(* IEC 61131-3 sources: SortJet_MasterSPS_Aufbau.fbsproj/Device.device.xml.v3^/Plc Logic.plclogic.xml.v3^/Application.application.xml.v3^/09_Station/Stationen/Faecherwagen [301-305]/0_Konfig, 5 files *)

(* ---- MK_Faecherwagen.gvl ---- *)
(* METADATA
{
	"v3Meta": {
		"objectGuid": "4f007b85-dd1b-4818-92fb-7451563e5cb0"
	}
}
*)
{attribute 'allow_unqualified_access'}
NAMESPACE MK_Faecherwagen
VAR_GLOBAL
  apgMKFaecherwagenstation : ARRAY[cERSTE_FAECHERWAGENSTATIONS_NR..cLETZTE_FAECHERWAGENSTATIONS_NR] OF Parameter_Station :=[
    (
     stStationsNummern         := (  NummerIntern    :=   301,                                 // Stationsnummer fuer das MMI und die Stationsangabe der Meldungen
                                     NummerExtern    :=  1301,                                 // Stationsnummer fuer Bedienermeldungen
                                     NummerSPS       :=   301 ),                               // Stationsnummer SPS-intern (Indizes)
      bDeaktivieren             := FALSE,                                                      // Station deaktiviert (keine Auftraege, keine Referenzfahrt)
      wMeldungsNummer           := 1400,                                                       // Basis-Meldungsnummer (WatchIO)
      eStationsTyp              := eFaecherwagen,                                              // Typ der Station
      eaAutomatikkreis          := [eAutomatikkreis_2],                                        // Automatikkreise, zu denen die Station gehoert
     // stStationsParameter
     // stSchnittstellendaten
     // stFremdanlage
     // stGlasdaten
      eaSicherheitskreis        := [eSicherheitskreis_1],                                      // Sicherheitskreise, in die die Station eingebunden ist
      // astSicherheitskreisTeilabschaltung
      eSystemcheckZyklus        := eSystemcheckZyklus_1,                                       // In welchem Zyklus des Systemchecks die Station geprueft wird
     // stStationsOptionen
      stStationsAufbau          := ( bAnschlag                     := FALSE,                   // Ausbaustufe: Ausrichtanschlaege
                                     bRolltor                      := TRUE,                    // Ausbaustufe Faecherwagen: Rolltor
                                     bKlemmzylinder                := FALSE,                   // Ausbaustufe Faecherwagen: Klemmzylinder fixiert den Oberrahmen beim Ein- und Ausschleusen
                                     bGreifer                      := [cANZAHL_WAENDE(FALSE)], // Shuttle: Greifer je Wand (Scheibe aus dem Faecherwagen ziehen bzw. hineinschieben)
                                     bRFID                         := TRUE,                    // RFID-Leser vorhanden
                                     bAGV                          := FALSE,                   // Ausbaustufe Faecherwagen: Betrieb mit AGV
                                     bGeblase                      := [ FALSE ],               // Ausbaustufe: Geblaese je Wand
                                     bGlastransport                := [ FALSE ],               // Ausbaustufe: Glastransport je Wand
                                     bKippen                       := [ FALSE ],               // Ausbaustufe: Kippen je Wand
                                     bTransportVerstellung         := [ FALSE ],               // Ausbaustufe Shuttle: Transport-/Dickenverstellung je Wand
                                     bWandverstellung              := [ FALSE ],               // Ausbaustufe Station: Wandverstellung je Wand
                                     bWandverstellungMotorisch     := FALSE,                   // Shuttle: Transport-/Wandverstellung mit Antrieb statt pneumatisch
                                     bRoellchenleiste              := [ FALSE ],               // Ausbaustufe Station: Roellchenleiste je Wand
                                     bHub                          := FALSE,                   // Ausbaustufe: Hub der Station
                                     bHubrahmen                    := FALSE,                   // Ausbaustufe: Hubrahmen (Riemen heben/senken)
                                     bDrehen                       := FALSE,                   // Ausbaustufe: Drehen
                                     bQuerachse                    := FALSE,                   // Ausbaustufe: Querachse
                                     bMessachse                    := FALSE,                   // Ausbaustufe: Messachse (Anlegetisch, Anlegewand)
                                     bDruckluft                    := FALSE,                   // Druckluftueberwachung vorhanden
                                     bSensorAuslauf                := FALSE,                   // Auslaufsensor vorhanden
                                     bSensorEinlauf                := FALSE,                   // Einlaufsensor vorhanden
                                     bSensorEinlaufStopp           := FALSE,                   // Shuttle: zusaetzlicher Stopp-Sensor am Einlauf (ohne: Einlaufsensor), Gegenstueck zum Auslauf-Stopp im Rueckwaertstransport
                                     bSensorAuslaufStopp           := FALSE,                   // Shuttle: zusaetzlicher Stopp-Sensor am Auslauf (ohne: Auslaufsensor), Verfahrfreigabe und Scheibe hat Shuttle verlassen
                                     bDurchlaufSperreZumNachfolger := FALSE,                   // Ausbaustufe: bewegliche Abschrankung zum Nachfolger
                                     bKippenSchuetz                := FALSE,                   // Kippen ueber Schuetz statt Umrichter
                                     bQuerfahrt                    := FALSE,                   // Ausbaustufe: Querfahrt
                                     bDurchgang                    := FALSE,                   // Station ist Teil eines Durchgangs (belegt = Oeffnen blockiert)
                                     bSlaveAntrieb                 := FALSE,                   // Glastransport mit Slave-Antrieb
                                     bKipparme                     := FALSE,                   // Ausbaustufe: Kipparme
                                     bMessachseAmEndeVomTisch      := FALSE,                   // Messachse am Ende des Tisches (Hoehenfehler fragt den Bediener)
                                     bDLSSchmiersystem             := FALSE,                   // Zentralschmierung DLS vorhanden
                                     bGlastransportSlaveVorhanden  := FALSE,                   // Glastransport mit Slave-Antrieb (Meldungen/Ueberwachung Slave)
                                     wHydraulikstation             := cHYDRAULIKSTATION_1      // Faecherwagen Hydraulik: zugeordnete Hydraulikstation (cHYDRAULIKSTATION_x), 0 = keine
                                    )
     // astShuttleAnhaltenQuellen
    ),
    (
     stStationsNummern         := (  NummerIntern    :=   302,                                 // Stationsnummer fuer das MMI und die Stationsangabe der Meldungen
                                     NummerExtern    :=  1302,                                 // Stationsnummer fuer Bedienermeldungen
                                     NummerSPS       :=   302 ),                               // Stationsnummer SPS-intern (Indizes)
      bDeaktivieren             := FALSE,                                                      // Station deaktiviert (keine Auftraege, keine Referenzfahrt)
      wMeldungsNummer           := 1420,                                                       // Basis-Meldungsnummer (WatchIO)
      eStationsTyp              := eFaecherwagen,                                              // Typ der Station
      eaAutomatikkreis          := [eAutomatikkreis_2],                                        // Automatikkreise, zu denen die Station gehoert
     // stStationsParameter
     // stSchnittstellendaten
     // stFremdanlage
     // stGlasdaten
      eaSicherheitskreis        := [eSicherheitskreis_1],                                      // Sicherheitskreise, in die die Station eingebunden ist
      // astSicherheitskreisTeilabschaltung
      eSystemcheckZyklus        := eSystemcheckZyklus_1,                                       // In welchem Zyklus des Systemchecks die Station geprueft wird
     // stStationsOptionen
      stStationsAufbau          := ( bAnschlag                     := FALSE,                   // Ausbaustufe: Ausrichtanschlaege
                                     bRolltor                      := TRUE,                    // Ausbaustufe Faecherwagen: Rolltor
                                     bKlemmzylinder                := FALSE,                   // Ausbaustufe Faecherwagen: Klemmzylinder fixiert den Oberrahmen beim Ein- und Ausschleusen
                                     bGreifer                      := [cANZAHL_WAENDE(FALSE)], // Shuttle: Greifer je Wand (Scheibe aus dem Faecherwagen ziehen bzw. hineinschieben)
                                     bRFID                         := TRUE,                    // RFID-Leser vorhanden
                                     bAGV                          := FALSE,                   // Ausbaustufe Faecherwagen: Betrieb mit AGV
                                     bGeblase                      := [ FALSE ],               // Ausbaustufe: Geblaese je Wand
                                     bGlastransport                := [ FALSE ],               // Ausbaustufe: Glastransport je Wand
                                     bKippen                       := [ FALSE ],               // Ausbaustufe: Kippen je Wand
                                     bTransportVerstellung         := [ FALSE ],               // Ausbaustufe Shuttle: Transport-/Dickenverstellung je Wand
                                     bWandverstellung              := [ FALSE ],               // Ausbaustufe Station: Wandverstellung je Wand
                                     bWandverstellungMotorisch     := FALSE,                   // Shuttle: Transport-/Wandverstellung mit Antrieb statt pneumatisch
                                     bRoellchenleiste              := [ FALSE ],               // Ausbaustufe Station: Roellchenleiste je Wand
                                     bHub                          := FALSE,                   // Ausbaustufe: Hub der Station
                                     bHubrahmen                    := FALSE,                   // Ausbaustufe: Hubrahmen (Riemen heben/senken)
                                     bDrehen                       := FALSE,                   // Ausbaustufe: Drehen
                                     bQuerachse                    := FALSE,                   // Ausbaustufe: Querachse
                                     bMessachse                    := FALSE,                   // Ausbaustufe: Messachse (Anlegetisch, Anlegewand)
                                     bDruckluft                    := FALSE,                   // Druckluftueberwachung vorhanden
                                     bSensorAuslauf                := FALSE,                   // Auslaufsensor vorhanden
                                     bSensorEinlauf                := FALSE,                   // Einlaufsensor vorhanden
                                     bSensorEinlaufStopp           := FALSE,                   // Shuttle: zusaetzlicher Stopp-Sensor am Einlauf (ohne: Einlaufsensor), Gegenstueck zum Auslauf-Stopp im Rueckwaertstransport
                                     bSensorAuslaufStopp           := FALSE,                   // Shuttle: zusaetzlicher Stopp-Sensor am Auslauf (ohne: Auslaufsensor), Verfahrfreigabe und Scheibe hat Shuttle verlassen
                                     bDurchlaufSperreZumNachfolger := FALSE,                   // Ausbaustufe: bewegliche Abschrankung zum Nachfolger
                                     bKippenSchuetz                := FALSE,                   // Kippen ueber Schuetz statt Umrichter
                                     bQuerfahrt                    := FALSE,                   // Ausbaustufe: Querfahrt
                                     bDurchgang                    := FALSE,                   // Station ist Teil eines Durchgangs (belegt = Oeffnen blockiert)
                                     bSlaveAntrieb                 := FALSE,                   // Glastransport mit Slave-Antrieb
                                     bKipparme                     := FALSE,                   // Ausbaustufe: Kipparme
                                     bMessachseAmEndeVomTisch      := FALSE,                   // Messachse am Ende des Tisches (Hoehenfehler fragt den Bediener)
                                     bDLSSchmiersystem             := FALSE,                   // Zentralschmierung DLS vorhanden
                                     bGlastransportSlaveVorhanden  := FALSE,                   // Glastransport mit Slave-Antrieb (Meldungen/Ueberwachung Slave)
                                     wHydraulikstation             := cHYDRAULIKSTATION_1      // Faecherwagen Hydraulik: zugeordnete Hydraulikstation (cHYDRAULIKSTATION_x), 0 = keine
                                    )
     // astShuttleAnhaltenQuellen
    ),
    (
     stStationsNummern         := (  NummerIntern    :=   303,                                 // Stationsnummer fuer das MMI und die Stationsangabe der Meldungen
                                     NummerExtern    :=  1303,                                 // Stationsnummer fuer Bedienermeldungen
                                     NummerSPS       :=   303 ),                               // Stationsnummer SPS-intern (Indizes)
      bDeaktivieren             := FALSE,                                                      // Station deaktiviert (keine Auftraege, keine Referenzfahrt)
      wMeldungsNummer           := 1440,                                                       // Basis-Meldungsnummer (WatchIO)
      eStationsTyp              := eFaecherwagen,                                              // Typ der Station
      eaAutomatikkreis          := [eAutomatikkreis_2],                                        // Automatikkreise, zu denen die Station gehoert
     // stStationsParameter
     // stSchnittstellendaten
     // stFremdanlage
     // stGlasdaten
      eaSicherheitskreis        := [eSicherheitskreis_1],                                      // Sicherheitskreise, in die die Station eingebunden ist
      // astSicherheitskreisTeilabschaltung
      eSystemcheckZyklus        := eSystemcheckZyklus_1,                                       // In welchem Zyklus des Systemchecks die Station geprueft wird
     // stStationsOptionen
      stStationsAufbau          := ( bAnschlag                     := FALSE,                   // Ausbaustufe: Ausrichtanschlaege
                                     bRolltor                      := TRUE,                    // Ausbaustufe Faecherwagen: Rolltor
                                     bKlemmzylinder                := FALSE,                   // Ausbaustufe Faecherwagen: Klemmzylinder fixiert den Oberrahmen beim Ein- und Ausschleusen
                                     bGreifer                      := [cANZAHL_WAENDE(FALSE)], // Shuttle: Greifer je Wand (Scheibe aus dem Faecherwagen ziehen bzw. hineinschieben)
                                     bRFID                         := TRUE,                    // RFID-Leser vorhanden
                                     bAGV                          := FALSE,                   // Ausbaustufe Faecherwagen: Betrieb mit AGV
                                     bGeblase                      := [ FALSE ],               // Ausbaustufe: Geblaese je Wand
                                     bGlastransport                := [ FALSE ],               // Ausbaustufe: Glastransport je Wand
                                     bKippen                       := [ FALSE ],               // Ausbaustufe: Kippen je Wand
                                     bTransportVerstellung         := [ FALSE ],               // Ausbaustufe Shuttle: Transport-/Dickenverstellung je Wand
                                     bWandverstellung              := [ FALSE ],               // Ausbaustufe Station: Wandverstellung je Wand
                                     bWandverstellungMotorisch     := FALSE,                   // Shuttle: Transport-/Wandverstellung mit Antrieb statt pneumatisch
                                     bRoellchenleiste              := [ FALSE ],               // Ausbaustufe Station: Roellchenleiste je Wand
                                     bHub                          := FALSE,                   // Ausbaustufe: Hub der Station
                                     bHubrahmen                    := FALSE,                   // Ausbaustufe: Hubrahmen (Riemen heben/senken)
                                     bDrehen                       := FALSE,                   // Ausbaustufe: Drehen
                                     bQuerachse                    := FALSE,                   // Ausbaustufe: Querachse
                                     bMessachse                    := FALSE,                   // Ausbaustufe: Messachse (Anlegetisch, Anlegewand)
                                     bDruckluft                    := FALSE,                   // Druckluftueberwachung vorhanden
                                     bSensorAuslauf                := FALSE,                   // Auslaufsensor vorhanden
                                     bSensorEinlauf                := FALSE,                   // Einlaufsensor vorhanden
                                     bSensorEinlaufStopp           := FALSE,                   // Shuttle: zusaetzlicher Stopp-Sensor am Einlauf (ohne: Einlaufsensor), Gegenstueck zum Auslauf-Stopp im Rueckwaertstransport
                                     bSensorAuslaufStopp           := FALSE,                   // Shuttle: zusaetzlicher Stopp-Sensor am Auslauf (ohne: Auslaufsensor), Verfahrfreigabe und Scheibe hat Shuttle verlassen
                                     bDurchlaufSperreZumNachfolger := FALSE,                   // Ausbaustufe: bewegliche Abschrankung zum Nachfolger
                                     bKippenSchuetz                := FALSE,                   // Kippen ueber Schuetz statt Umrichter
                                     bQuerfahrt                    := FALSE,                   // Ausbaustufe: Querfahrt
                                     bDurchgang                    := FALSE,                   // Station ist Teil eines Durchgangs (belegt = Oeffnen blockiert)
                                     bSlaveAntrieb                 := FALSE,                   // Glastransport mit Slave-Antrieb
                                     bKipparme                     := FALSE,                   // Ausbaustufe: Kipparme
                                     bMessachseAmEndeVomTisch      := FALSE,                   // Messachse am Ende des Tisches (Hoehenfehler fragt den Bediener)
                                     bDLSSchmiersystem             := FALSE,                   // Zentralschmierung DLS vorhanden
                                     bGlastransportSlaveVorhanden  := FALSE,                   // Glastransport mit Slave-Antrieb (Meldungen/Ueberwachung Slave)
                                     wHydraulikstation             := cHYDRAULIKSTATION_1      // Faecherwagen Hydraulik: zugeordnete Hydraulikstation (cHYDRAULIKSTATION_x), 0 = keine
                                    )
     // astShuttleAnhaltenQuellen
    ),
    (
     stStationsNummern         := (  NummerIntern    :=   304,                                 // Stationsnummer fuer das MMI und die Stationsangabe der Meldungen
                                     NummerExtern    :=  1304,                                 // Stationsnummer fuer Bedienermeldungen
                                     NummerSPS       :=   304 ),                               // Stationsnummer SPS-intern (Indizes)
      bDeaktivieren             := FALSE,                                                      // Station deaktiviert (keine Auftraege, keine Referenzfahrt)
      wMeldungsNummer           := 1460,                                                       // Basis-Meldungsnummer (WatchIO)
      eStationsTyp              := eFaecherwagen,                                              // Typ der Station
      eaAutomatikkreis          := [eAutomatikkreis_2],                                        // Automatikkreise, zu denen die Station gehoert
     // stStationsParameter
     // stSchnittstellendaten
     // stFremdanlage
     // stGlasdaten
      eaSicherheitskreis        := [eSicherheitskreis_1],                                      // Sicherheitskreise, in die die Station eingebunden ist
      // astSicherheitskreisTeilabschaltung
      eSystemcheckZyklus        := eSystemcheckZyklus_1,                                       // In welchem Zyklus des Systemchecks die Station geprueft wird
     // stStationsOptionen
      stStationsAufbau          := ( bAnschlag                     := FALSE,                   // Ausbaustufe: Ausrichtanschlaege
                                     bRolltor                      := TRUE,                    // Ausbaustufe Faecherwagen: Rolltor
                                     bKlemmzylinder                := FALSE,                   // Ausbaustufe Faecherwagen: Klemmzylinder fixiert den Oberrahmen beim Ein- und Ausschleusen
                                     bGreifer                      := [cANZAHL_WAENDE(FALSE)], // Shuttle: Greifer je Wand (Scheibe aus dem Faecherwagen ziehen bzw. hineinschieben)
                                     bRFID                         := TRUE,                    // RFID-Leser vorhanden
                                     bAGV                          := FALSE,                   // Ausbaustufe Faecherwagen: Betrieb mit AGV
                                     bGeblase                      := [ FALSE ],               // Ausbaustufe: Geblaese je Wand
                                     bGlastransport                := [ FALSE ],               // Ausbaustufe: Glastransport je Wand
                                     bKippen                       := [ FALSE ],               // Ausbaustufe: Kippen je Wand
                                     bTransportVerstellung         := [ FALSE ],               // Ausbaustufe Shuttle: Transport-/Dickenverstellung je Wand
                                     bWandverstellung              := [ FALSE ],               // Ausbaustufe Station: Wandverstellung je Wand
                                     bWandverstellungMotorisch     := FALSE,                   // Shuttle: Transport-/Wandverstellung mit Antrieb statt pneumatisch
                                     bRoellchenleiste              := [ FALSE ],               // Ausbaustufe Station: Roellchenleiste je Wand
                                     bHub                          := FALSE,                   // Ausbaustufe: Hub der Station
                                     bHubrahmen                    := FALSE,                   // Ausbaustufe: Hubrahmen (Riemen heben/senken)
                                     bDrehen                       := FALSE,                   // Ausbaustufe: Drehen
                                     bQuerachse                    := FALSE,                   // Ausbaustufe: Querachse
                                     bMessachse                    := FALSE,                   // Ausbaustufe: Messachse (Anlegetisch, Anlegewand)
                                     bDruckluft                    := FALSE,                   // Druckluftueberwachung vorhanden
                                     bSensorAuslauf                := FALSE,                   // Auslaufsensor vorhanden
                                     bSensorEinlauf                := FALSE,                   // Einlaufsensor vorhanden
                                     bSensorEinlaufStopp           := FALSE,                   // Shuttle: zusaetzlicher Stopp-Sensor am Einlauf (ohne: Einlaufsensor), Gegenstueck zum Auslauf-Stopp im Rueckwaertstransport
                                     bSensorAuslaufStopp           := FALSE,                   // Shuttle: zusaetzlicher Stopp-Sensor am Auslauf (ohne: Auslaufsensor), Verfahrfreigabe und Scheibe hat Shuttle verlassen
                                     bDurchlaufSperreZumNachfolger := FALSE,                   // Ausbaustufe: bewegliche Abschrankung zum Nachfolger
                                     bKippenSchuetz                := FALSE,                   // Kippen ueber Schuetz statt Umrichter
                                     bQuerfahrt                    := FALSE,                   // Ausbaustufe: Querfahrt
                                     bDurchgang                    := FALSE,                   // Station ist Teil eines Durchgangs (belegt = Oeffnen blockiert)
                                     bSlaveAntrieb                 := FALSE,                   // Glastransport mit Slave-Antrieb
                                     bKipparme                     := FALSE,                   // Ausbaustufe: Kipparme
                                     bMessachseAmEndeVomTisch      := FALSE,                   // Messachse am Ende des Tisches (Hoehenfehler fragt den Bediener)
                                     bDLSSchmiersystem             := FALSE,                   // Zentralschmierung DLS vorhanden
                                     bGlastransportSlaveVorhanden  := FALSE,                   // Glastransport mit Slave-Antrieb (Meldungen/Ueberwachung Slave)
                                     wHydraulikstation             := cHYDRAULIKSTATION_1      // Faecherwagen Hydraulik: zugeordnete Hydraulikstation (cHYDRAULIKSTATION_x), 0 = keine
                                    )
     // astShuttleAnhaltenQuellen
    ),
    (
     stStationsNummern         := (  NummerIntern    :=   305,                                 // Stationsnummer fuer das MMI und die Stationsangabe der Meldungen
                                     NummerExtern    :=  1305,                                 // Stationsnummer fuer Bedienermeldungen
                                     NummerSPS       :=   305 ),                               // Stationsnummer SPS-intern (Indizes)
      bDeaktivieren             := FALSE,                                                      // Station deaktiviert (keine Auftraege, keine Referenzfahrt)
      wMeldungsNummer           := 1480,                                                       // Basis-Meldungsnummer (WatchIO)
      eStationsTyp              := eFaecherwagen,                                              // Typ der Station
      eaAutomatikkreis          := [eAutomatikkreis_2],                                        // Automatikkreise, zu denen die Station gehoert
     // stStationsParameter
     // stSchnittstellendaten
     // stFremdanlage
     // stGlasdaten
      eaSicherheitskreis        := [eSicherheitskreis_1],                                      // Sicherheitskreise, in die die Station eingebunden ist
      // astSicherheitskreisTeilabschaltung
      eSystemcheckZyklus        := eSystemcheckZyklus_1,                                       // In welchem Zyklus des Systemchecks die Station geprueft wird
     // stStationsOptionen
      stStationsAufbau          := ( bAnschlag                     := FALSE,                   // Ausbaustufe: Ausrichtanschlaege
                                     bRolltor                      := TRUE,                    // Ausbaustufe Faecherwagen: Rolltor
                                     bKlemmzylinder                := FALSE,                   // Ausbaustufe Faecherwagen: Klemmzylinder fixiert den Oberrahmen beim Ein- und Ausschleusen
                                     bGreifer                      := [cANZAHL_WAENDE(FALSE)], // Shuttle: Greifer je Wand (Scheibe aus dem Faecherwagen ziehen bzw. hineinschieben)
                                     bRFID                         := TRUE,                    // RFID-Leser vorhanden
                                     bAGV                          := FALSE,                   // Ausbaustufe Faecherwagen: Betrieb mit AGV
                                     bGeblase                      := [ FALSE ],               // Ausbaustufe: Geblaese je Wand
                                     bGlastransport                := [ FALSE ],               // Ausbaustufe: Glastransport je Wand
                                     bKippen                       := [ FALSE ],               // Ausbaustufe: Kippen je Wand
                                     bTransportVerstellung         := [ FALSE ],               // Ausbaustufe Shuttle: Transport-/Dickenverstellung je Wand
                                     bWandverstellung              := [ FALSE ],               // Ausbaustufe Station: Wandverstellung je Wand
                                     bWandverstellungMotorisch     := FALSE,                   // Shuttle: Transport-/Wandverstellung mit Antrieb statt pneumatisch
                                     bRoellchenleiste              := [ FALSE ],               // Ausbaustufe Station: Roellchenleiste je Wand
                                     bHub                          := FALSE,                   // Ausbaustufe: Hub der Station
                                     bHubrahmen                    := FALSE,                   // Ausbaustufe: Hubrahmen (Riemen heben/senken)
                                     bDrehen                       := FALSE,                   // Ausbaustufe: Drehen
                                     bQuerachse                    := FALSE,                   // Ausbaustufe: Querachse
                                     bMessachse                    := FALSE,                   // Ausbaustufe: Messachse (Anlegetisch, Anlegewand)
                                     bDruckluft                    := FALSE,                   // Druckluftueberwachung vorhanden
                                     bSensorAuslauf                := FALSE,                   // Auslaufsensor vorhanden
                                     bSensorEinlauf                := FALSE,                   // Einlaufsensor vorhanden
                                     bSensorEinlaufStopp           := FALSE,                   // Shuttle: zusaetzlicher Stopp-Sensor am Einlauf (ohne: Einlaufsensor), Gegenstueck zum Auslauf-Stopp im Rueckwaertstransport
                                     bSensorAuslaufStopp           := FALSE,                   // Shuttle: zusaetzlicher Stopp-Sensor am Auslauf (ohne: Auslaufsensor), Verfahrfreigabe und Scheibe hat Shuttle verlassen
                                     bDurchlaufSperreZumNachfolger := FALSE,                   // Ausbaustufe: bewegliche Abschrankung zum Nachfolger
                                     bKippenSchuetz                := FALSE,                   // Kippen ueber Schuetz statt Umrichter
                                     bQuerfahrt                    := FALSE,                   // Ausbaustufe: Querfahrt
                                     bDurchgang                    := FALSE,                   // Station ist Teil eines Durchgangs (belegt = Oeffnen blockiert)
                                     bSlaveAntrieb                 := FALSE,                   // Glastransport mit Slave-Antrieb
                                     bKipparme                     := FALSE,                   // Ausbaustufe: Kipparme
                                     bMessachseAmEndeVomTisch      := FALSE,                   // Messachse am Ende des Tisches (Hoehenfehler fragt den Bediener)
                                     bDLSSchmiersystem             := FALSE,                   // Zentralschmierung DLS vorhanden
                                     bGlastransportSlaveVorhanden  := FALSE,                   // Glastransport mit Slave-Antrieb (Meldungen/Ueberwachung Slave)
                                     wHydraulikstation             := cHYDRAULIKSTATION_1      // Faecherwagen Hydraulik: zugeordnete Hydraulikstation (cHYDRAULIKSTATION_x), 0 = keine
                                    )
     // astShuttleAnhaltenQuellen
    )];

END_VAR
END_NAMESPACE

(* ---- MK_Hydraulikstation.gvl ---- *)
(* METADATA
{
	"v3Meta": {
		"objectGuid": "ffb6da21-2d1f-4f73-afc8-e550ef19dd3a"
	}
}
*)
{attribute 'allow_unqualified_access'}
NAMESPACE MK_Hydraulikstation
VAR_GLOBAL
  // Hydraulikaggregate der Faecherwagenstationen (Variante Hydraulik)
  // Zuordnung Faecherwagenstation -> Hydraulikstation: MK stStationsAufbau.wHydraulikstation der Faecherwagenstation
  apgMKHydraulikstation : ARRAY[cERSTE_HYDRAULIKSTATIONS_NR..cLETZTE_HYDRAULIKSTATIONS_NR] OF Parameter_Hydraulikstation :=[
    (
      bDeaktivieren                   := TRUE, // Station deaktiviert (keine Auftraege, keine Referenzfahrt)
      wMeldungsNummer                 := 2000, // WatchIO-Meldung Motorschutz Hydraulikaggregat
      wMaximaleAnzahlAktiverAuftraege := 1     // Max. gleichzeitige Ein-/Ausschleus-Auftraege der zugeordneten Stationen, 0 = unbegrenzt
    )];

END_VAR

END_NAMESPACE

(* ---- Konfiguration_FW_Basis.gvl ---- *)
(* METADATA
{
	"v3Meta": {
		"objectGuid": "7937dd0c-d972-4971-bda8-59bd0e2e5387"
	}
}
*)
{attribute 'allow_unqualified_access'}
NAMESPACE Konfiguration_FW_Basis
VAR_CONFIG

//-------------------------------------------------------------------------------------------------
// KONFIGURATION: BASISKOMPONENTEN
//-------------------------------------------------------------------------------------------------

  // ------------------------------------ HARDWARE EINGAENGE ---------------------------------------
  // EINGAENGE: Hydraulikstation 1 (cHYDRAULIKSTATION_1)
  Globale_Bausteine.aHydraulikstation[1].in_bMotorschuetz_Hydraulikkreislauf_OK              AT %MX1.1    : BOOL; // OPTION

  // ------------------------------------ HARDWARE AUSGAENGE ---------------------------------------
  // AUSGAENGE: Hydraulikstation 1 (cHYDRAULIKSTATION_1)
  Globale_Bausteine.aHydraulikstation[1].out_bHydraulikkreislauf_MotorEin                    AT %MX3000.0 : BOOL; // OPTION
  Globale_Bausteine.aHydraulikstation[1].out_bHydraulikkreislauf_UmlaufventilAuf             AT %MX3000.1 : BOOL; // OPTION

Globale_Bausteine.aFaecherwagenstation[301].out_bRolltorAb                                   AT %QX11.0  : BOOL; // IO-L - Rolltor 301 schliessen
Globale_Bausteine.aFaecherwagenstation[301].out_bRolltorAuf                                  AT %QX11.1  : BOOL; // IO-L - Rolltor 301 oeffnen
Globale_Bausteine.aFaecherwagenstation[302].out_bRolltorAb                                   AT %QX11.2  : BOOL; // IO-L - Rolltor 302 schliessen
Globale_Bausteine.aFaecherwagenstation[302].out_bRolltorAuf                                  AT %QX11.3  : BOOL; // IO-L - Rolltor 302 oeffnen
Globale_Bausteine.aFaecherwagenstation[303].out_bRolltorAb                                   AT %QX11.4  : BOOL; // IO-L - Rolltor 303 schliessen
Globale_Bausteine.aFaecherwagenstation[303].out_bRolltorAuf                                  AT %QX11.5  : BOOL; // IO-L - Rolltor 303 oeffnen
Globale_Bausteine.aFaecherwagenstation[304].out_bRolltorAb                                   AT %QX11.6   : BOOL; // IO-L - Rolltor 304 schliessen
Globale_Bausteine.aFaecherwagenstation[304].out_bRolltorAuf                                  AT %QX11.7   : BOOL; // IO-L - Rolltor 304 oeffnen
Globale_Bausteine.aFaecherwagenstation[305].out_bRolltorAb                                   AT %QX12.0   : BOOL; // IO-L - Rolltor 305 schliessen
Globale_Bausteine.aFaecherwagenstation[305].out_bRolltorAuf                                  AT %QX12.1   : BOOL; // IO-L - Rolltor 305 oeffnen

  // Rolltor oben (in_bNichtRolltorGeoeffnet), Sicherheitskreis und sichere Feldbox: im Geraetebaum gemappt

  // Varianten Einfach und Hydraulik: IOs je Station in Konfiguration_FW_Einfach bzw. Konfiguration_FW_Hydraulik

END_VAR

END_NAMESPACE

(* ---- Konfiguration_FW_Einfach.gvl ---- *)
(* METADATA
{
	"v3Meta": {
		"objectGuid": "02dda72b-1e55-4a9f-86bc-3e1987758175"
	}
}
*)
{attribute 'allow_unqualified_access'}
NAMESPACE Konfiguration_FW_Einfach
VAR_CONFIG

//-------------------------------------------------------------------------------------------------
// KONFIGURATION: FAECHERWAGENSTATIONEN VARIANTE EINFACH
// Nur verwenden, wenn aFaecherwagenstation (Globale_Bausteine) vom Typ Faecherwagenstation_Einfach_FB_V01_00_00 ist,
// sonst Attribut excludefrombuild setzen. Es darf immer nur eine Variante im Build sein.
// Arretierung (Gegenhalter) und Schleusen-Taster/-Leuchte liegen am IO-Link und sind im Geraetebaum gemappt.
// Faecherwagen vorhanden kommt aus der SLC (Interface_SLC, bpFaecherwagenVorhanden).
// Platzhalter: Eingaenge %MX1.0 (FALSE) / %MX1.1 (TRUE)
//-------------------------------------------------------------------------------------------------

  // ------------------------------------ STATION 301 ------------------------------------------------
  // EINGAENGE
  Globale_Bausteine.aFaecherwagenstation[301].in_bAbrollsicherungOK                             AT %IX0.1    : BOOL; // IO-L - Abrollsicherung OK (Sammelmeldung Versorgung FW1 Rolltore / Abrollsicherung OK)

  // ------------------------------------ STATION 302 ------------------------------------------------
  // EINGAENGE
  Globale_Bausteine.aFaecherwagenstation[302].in_bAbrollsicherungOK                             AT %IX0.1    : BOOL; // IO-L - Abrollsicherung OK (Sammelmeldung Versorgung FW1 Rolltore / Abrollsicherung OK)

  // ------------------------------------ STATION 303 ------------------------------------------------
  // EINGAENGE
  Globale_Bausteine.aFaecherwagenstation[303].in_bAbrollsicherungOK                             AT %IX0.1    : BOOL; // IO-L - Abrollsicherung OK (Sammelmeldung Versorgung FW1 Rolltore / Abrollsicherung OK)

  // ------------------------------------ STATION 304 ------------------------------------------------
  // EINGAENGE
  Globale_Bausteine.aFaecherwagenstation[304].in_bAbrollsicherungOK                             AT %IX0.1    : BOOL; // IO-L - Abrollsicherung OK (Sammelmeldung Versorgung FW1 Rolltore / Abrollsicherung OK)

  // ------------------------------------ STATION 305 ------------------------------------------------
  // EINGAENGE
  Globale_Bausteine.aFaecherwagenstation[305].in_bAbrollsicherungOK                             AT %IX0.1    : BOOL; // IO-L - Abrollsicherung OK (Sammelmeldung Versorgung FW1 Rolltore / Abrollsicherung OK)

END_VAR

END_NAMESPACE

(* ---- Konfiguration_FW_Hydraulik.gvl ---- *)
(* METADATA
{
	"v3Meta": {
		"objectGuid": "402b1ef0-d461-45b4-8faf-9d71f219f2c1"
	}
}
*)
{attribute 'excludefrombuild'}
{attribute 'allow_unqualified_access'}
NAMESPACE Konfiguration_FW_Hydraulik
VAR_CONFIG

//-------------------------------------------------------------------------------------------------
// KONFIGURATION: FAECHERWAGENSTATIONEN VARIANTE HYDRAULIK
// Nur verwenden, wenn aFaecherwagenstation (Globale_Bausteine) vom Typ Faecherwagenstation_Hydraulik_FB_V01_00_00 ist:
// dann Attribut excludefrombuild entfernen. Es darf immer nur eine Variante im Build sein.
// Platzhalter: Eingaenge %MX1.0 (FALSE) / %MX1.1 (TRUE), Ausgaenge je Station ab %MX<Station*10>.0
//-------------------------------------------------------------------------------------------------

  // ------------------------------------ STATION 301 ------------------------------------------------
  // EINGAENGE
  Globale_Bausteine.aFaecherwagenstation[301].in_bHubrahmenOben                                 AT %MX1.0    : BOOL; // OPTION - Hubrahmen oben 301, aus Schaltplan
  Globale_Bausteine.aFaecherwagenstation[301].in_bHubrahmenUnten                                AT %MX1.0    : BOOL; // OPTION - Hubrahmen unten 301, aus Schaltplan
  Globale_Bausteine.aFaecherwagenstation[301].in_bFaecherwagenVorne                             AT %MX1.0    : BOOL; // OPTION - Faecherwagen vorne 301, aus Schaltplan
  Globale_Bausteine.aFaecherwagenstation[301].in_bFaecherwagenHinten                            AT %MX1.0    : BOOL; // OPTION - Faecherwagen hinten 301, aus Schaltplan
  Globale_Bausteine.aFaecherwagenstation[301].in_bZentrierungOffen                              AT %MX1.0    : BOOL; // OPTION - Zentrierung offen 301, aus Schaltplan
  Globale_Bausteine.aFaecherwagenstation[301].in_bZentrierungGeschlossen                        AT %MX1.0    : BOOL; // OPTION - Zentrierung geschlossen 301, aus Schaltplan
  Globale_Bausteine.aFaecherwagenstation[301].in_bAnschlagOben                                  AT %MX1.0    : BOOL; // OPTION - Anschlag oben 301, aus Schaltplan
  Globale_Bausteine.aFaecherwagenstation[301].in_bAnschlagUnten                                 AT %MX1.0    : BOOL; // OPTION - Anschlag unten 301, aus Schaltplan
  Globale_Bausteine.aFaecherwagenstation[301].in_bAnschlagVorne                                 AT %MX1.0    : BOOL; // OPTION - OPTION AGV: Anschlag vorne 301, aus Schaltplan
  Globale_Bausteine.aFaecherwagenstation[301].in_bAnschlagHinten                                AT %MX1.0    : BOOL; // OPTION - OPTION AGV: Anschlag hinten 301, aus Schaltplan
  Globale_Bausteine.aFaecherwagenstation[301].in_bFWInAusrichtPosition                          AT %MX1.0    : BOOL; // OPTION - Faecherwagen in Ausrichtposition 301, aus Schaltplan
  Globale_Bausteine.aFaecherwagenstation[301].in_bMutingSensorLinks                             AT %MX1.0    : BOOL; // OPTION - Muting-Sensor links 301, aus Schaltplan
  Globale_Bausteine.aFaecherwagenstation[301].in_bMutingSensorRechts                            AT %MX1.0    : BOOL; // OPTION - Muting-Sensor rechts 301, aus Schaltplan
  Globale_Bausteine.aFaecherwagenstation[301].in_bStartSchleusen                                AT %MX1.0    : BOOL; // OPTION - Taster Ein-/Ausschleusen 301, aus Schaltplan
  Globale_Bausteine.aFaecherwagenstation[301].in_bSicherheitsrelaisOK                           AT %MX1.1    : BOOL; // OPTION - Sicherheitsrelais in Ordnung 301, aus Schaltplan
  Globale_Bausteine.aFaecherwagenstation[301].in_bAbrollsicherungOK                             AT %MX1.1    : BOOL; // OPTION - Abrollsicherung des Rolltors nicht ausgeloest 301, aus Schaltplan
  Globale_Bausteine.aFaecherwagenstation[301].in_bRFID_DataValid                                AT %MX1.0    : BOOL; // OPTION - RFID Daten gueltig 301, aus Schaltplan
  Globale_Bausteine.aFaecherwagenstation[301].in_bRFID_NR1                                      AT %MX1.0    : BOOL; // OPTION - RFID Bit 1 301, aus Schaltplan
  Globale_Bausteine.aFaecherwagenstation[301].in_bRFID_NR2                                      AT %MX1.0    : BOOL; // OPTION - RFID Bit 2 301, aus Schaltplan
  Globale_Bausteine.aFaecherwagenstation[301].in_bRFID_NR3                                      AT %MX1.0    : BOOL; // OPTION - RFID Bit 3 301, aus Schaltplan
  Globale_Bausteine.aFaecherwagenstation[301].in_bRFID_NR4                                      AT %MX1.0    : BOOL; // OPTION - RFID Bit 4 301, aus Schaltplan
  Globale_Bausteine.aFaecherwagenstation[301].in_bRFID_NR5                                      AT %MX1.0    : BOOL; // OPTION - RFID Bit 5 301, aus Schaltplan
  Globale_Bausteine.aFaecherwagenstation[301].in_bRFID_NR6                                      AT %MX1.0    : BOOL; // OPTION - RFID Bit 6 301, aus Schaltplan
  Globale_Bausteine.aFaecherwagenstation[301].in_bRFID_NR7                                      AT %MX1.0    : BOOL; // OPTION - RFID Bit 7 301, aus Schaltplan
  Globale_Bausteine.aFaecherwagenstation[301].in_bRFID_NR8                                      AT %MX1.0    : BOOL; // OPTION - RFID Bit 8 301, aus Schaltplan
  // AUSGAENGE
  Globale_Bausteine.aFaecherwagenstation[301].out_bHubrahmenHeben                               AT %MX3010.0 : BOOL; // OPTION - Hubrahmen heben 301, aus Schaltplan
  Globale_Bausteine.aFaecherwagenstation[301].out_bHubrahmenSenken                              AT %MX3010.1 : BOOL; // OPTION - Hubrahmen senken 301, aus Schaltplan
  Globale_Bausteine.aFaecherwagenstation[301].out_bFaecherwagenVor                              AT %MX3010.2 : BOOL; // OPTION - Faecherwagen vor 301, aus Schaltplan
  Globale_Bausteine.aFaecherwagenstation[301].out_bFaecherwagenZurueck                          AT %MX3010.3 : BOOL; // OPTION - Faecherwagen zurueck 301, aus Schaltplan
  Globale_Bausteine.aFaecherwagenstation[301].out_bZentrierungOeffnen                           AT %MX3010.4 : BOOL; // OPTION - Zentrierung oeffnen 301, aus Schaltplan
  Globale_Bausteine.aFaecherwagenstation[301].out_bZentrierungSchliessen                        AT %MX3010.5 : BOOL; // OPTION - Zentrierung schliessen 301, aus Schaltplan
  Globale_Bausteine.aFaecherwagenstation[301].out_bAnschlagAuf                                  AT %MX3010.6 : BOOL; // OPTION - Anschlag auf 301, aus Schaltplan
  Globale_Bausteine.aFaecherwagenstation[301].out_bAnschlagAb                                   AT %MX3010.7 : BOOL; // OPTION - Anschlag ab 301, aus Schaltplan
  Globale_Bausteine.aFaecherwagenstation[301].out_bAnschlagVor                                  AT %MX3011.0 : BOOL; // OPTION - OPTION AGV: Anschlag vor 301, aus Schaltplan
  Globale_Bausteine.aFaecherwagenstation[301].out_bAnschlagZurueck                              AT %MX3011.1 : BOOL; // OPTION - OPTION AGV: Anschlag zurueck 301, aus Schaltplan
  Globale_Bausteine.aFaecherwagenstation[301].out_bFreigabeSchleusen                            AT %MX3011.2 : BOOL; // OPTION - Leuchte im Taster Ein-/Ausschleusen 301, aus Schaltplan
  Globale_Bausteine.aFaecherwagenstation[301].out_bMutingSensorReset                            AT %MX3011.3 : BOOL; // OPTION - Reset Muting-Sensoren 301, aus Schaltplan
  Globale_Bausteine.aFaecherwagenstation[301].out_bResetSicherheitsrelais                       AT %MX3011.4 : BOOL; // OPTION - Reset Sicherheitsrelais 301, aus Schaltplan

  // ------------------------------------ STATION 302 ------------------------------------------------
  // EINGAENGE
  Globale_Bausteine.aFaecherwagenstation[302].in_bHubrahmenOben                                 AT %MX1.0    : BOOL; // OPTION - Hubrahmen oben 302, aus Schaltplan
  Globale_Bausteine.aFaecherwagenstation[302].in_bHubrahmenUnten                                AT %MX1.0    : BOOL; // OPTION - Hubrahmen unten 302, aus Schaltplan
  Globale_Bausteine.aFaecherwagenstation[302].in_bFaecherwagenVorne                             AT %MX1.0    : BOOL; // OPTION - Faecherwagen vorne 302, aus Schaltplan
  Globale_Bausteine.aFaecherwagenstation[302].in_bFaecherwagenHinten                            AT %MX1.0    : BOOL; // OPTION - Faecherwagen hinten 302, aus Schaltplan
  Globale_Bausteine.aFaecherwagenstation[302].in_bZentrierungOffen                              AT %MX1.0    : BOOL; // OPTION - Zentrierung offen 302, aus Schaltplan
  Globale_Bausteine.aFaecherwagenstation[302].in_bZentrierungGeschlossen                        AT %MX1.0    : BOOL; // OPTION - Zentrierung geschlossen 302, aus Schaltplan
  Globale_Bausteine.aFaecherwagenstation[302].in_bAnschlagOben                                  AT %MX1.0    : BOOL; // OPTION - Anschlag oben 302, aus Schaltplan
  Globale_Bausteine.aFaecherwagenstation[302].in_bAnschlagUnten                                 AT %MX1.0    : BOOL; // OPTION - Anschlag unten 302, aus Schaltplan
  Globale_Bausteine.aFaecherwagenstation[302].in_bAnschlagVorne                                 AT %MX1.0    : BOOL; // OPTION - OPTION AGV: Anschlag vorne 302, aus Schaltplan
  Globale_Bausteine.aFaecherwagenstation[302].in_bAnschlagHinten                                AT %MX1.0    : BOOL; // OPTION - OPTION AGV: Anschlag hinten 302, aus Schaltplan
  Globale_Bausteine.aFaecherwagenstation[302].in_bFWInAusrichtPosition                          AT %MX1.0    : BOOL; // OPTION - Faecherwagen in Ausrichtposition 302, aus Schaltplan
  Globale_Bausteine.aFaecherwagenstation[302].in_bMutingSensorLinks                             AT %MX1.0    : BOOL; // OPTION - Muting-Sensor links 302, aus Schaltplan
  Globale_Bausteine.aFaecherwagenstation[302].in_bMutingSensorRechts                            AT %MX1.0    : BOOL; // OPTION - Muting-Sensor rechts 302, aus Schaltplan
  Globale_Bausteine.aFaecherwagenstation[302].in_bStartSchleusen                                AT %MX1.0    : BOOL; // OPTION - Taster Ein-/Ausschleusen 302, aus Schaltplan
  Globale_Bausteine.aFaecherwagenstation[302].in_bSicherheitsrelaisOK                           AT %MX1.1    : BOOL; // OPTION - Sicherheitsrelais in Ordnung 302, aus Schaltplan
  Globale_Bausteine.aFaecherwagenstation[302].in_bAbrollsicherungOK                             AT %MX1.1    : BOOL; // OPTION - Abrollsicherung des Rolltors nicht ausgeloest 302, aus Schaltplan
  Globale_Bausteine.aFaecherwagenstation[302].in_bRFID_DataValid                                AT %MX1.0    : BOOL; // OPTION - RFID Daten gueltig 302, aus Schaltplan
  Globale_Bausteine.aFaecherwagenstation[302].in_bRFID_NR1                                      AT %MX1.0    : BOOL; // OPTION - RFID Bit 1 302, aus Schaltplan
  Globale_Bausteine.aFaecherwagenstation[302].in_bRFID_NR2                                      AT %MX1.0    : BOOL; // OPTION - RFID Bit 2 302, aus Schaltplan
  Globale_Bausteine.aFaecherwagenstation[302].in_bRFID_NR3                                      AT %MX1.0    : BOOL; // OPTION - RFID Bit 3 302, aus Schaltplan
  Globale_Bausteine.aFaecherwagenstation[302].in_bRFID_NR4                                      AT %MX1.0    : BOOL; // OPTION - RFID Bit 4 302, aus Schaltplan
  Globale_Bausteine.aFaecherwagenstation[302].in_bRFID_NR5                                      AT %MX1.0    : BOOL; // OPTION - RFID Bit 5 302, aus Schaltplan
  Globale_Bausteine.aFaecherwagenstation[302].in_bRFID_NR6                                      AT %MX1.0    : BOOL; // OPTION - RFID Bit 6 302, aus Schaltplan
  Globale_Bausteine.aFaecherwagenstation[302].in_bRFID_NR7                                      AT %MX1.0    : BOOL; // OPTION - RFID Bit 7 302, aus Schaltplan
  Globale_Bausteine.aFaecherwagenstation[302].in_bRFID_NR8                                      AT %MX1.0    : BOOL; // OPTION - RFID Bit 8 302, aus Schaltplan
  // AUSGAENGE
  Globale_Bausteine.aFaecherwagenstation[302].out_bHubrahmenHeben                               AT %MX3020.0 : BOOL; // OPTION - Hubrahmen heben 302, aus Schaltplan
  Globale_Bausteine.aFaecherwagenstation[302].out_bHubrahmenSenken                              AT %MX3020.1 : BOOL; // OPTION - Hubrahmen senken 302, aus Schaltplan
  Globale_Bausteine.aFaecherwagenstation[302].out_bFaecherwagenVor                              AT %MX3020.2 : BOOL; // OPTION - Faecherwagen vor 302, aus Schaltplan
  Globale_Bausteine.aFaecherwagenstation[302].out_bFaecherwagenZurueck                          AT %MX3020.3 : BOOL; // OPTION - Faecherwagen zurueck 302, aus Schaltplan
  Globale_Bausteine.aFaecherwagenstation[302].out_bZentrierungOeffnen                           AT %MX3020.4 : BOOL; // OPTION - Zentrierung oeffnen 302, aus Schaltplan
  Globale_Bausteine.aFaecherwagenstation[302].out_bZentrierungSchliessen                        AT %MX3020.5 : BOOL; // OPTION - Zentrierung schliessen 302, aus Schaltplan
  Globale_Bausteine.aFaecherwagenstation[302].out_bAnschlagAuf                                  AT %MX3020.6 : BOOL; // OPTION - Anschlag auf 302, aus Schaltplan
  Globale_Bausteine.aFaecherwagenstation[302].out_bAnschlagAb                                   AT %MX3020.7 : BOOL; // OPTION - Anschlag ab 302, aus Schaltplan
  Globale_Bausteine.aFaecherwagenstation[302].out_bAnschlagVor                                  AT %MX3021.0 : BOOL; // OPTION - OPTION AGV: Anschlag vor 302, aus Schaltplan
  Globale_Bausteine.aFaecherwagenstation[302].out_bAnschlagZurueck                              AT %MX3021.1 : BOOL; // OPTION - OPTION AGV: Anschlag zurueck 302, aus Schaltplan
  Globale_Bausteine.aFaecherwagenstation[302].out_bFreigabeSchleusen                            AT %MX3021.2 : BOOL; // OPTION - Leuchte im Taster Ein-/Ausschleusen 302, aus Schaltplan
  Globale_Bausteine.aFaecherwagenstation[302].out_bMutingSensorReset                            AT %MX3021.3 : BOOL; // OPTION - Reset Muting-Sensoren 302, aus Schaltplan
  Globale_Bausteine.aFaecherwagenstation[302].out_bResetSicherheitsrelais                       AT %MX3021.4 : BOOL; // OPTION - Reset Sicherheitsrelais 302, aus Schaltplan

  // ------------------------------------ STATION 303 ------------------------------------------------
  // EINGAENGE
  Globale_Bausteine.aFaecherwagenstation[303].in_bHubrahmenOben                                 AT %MX1.0    : BOOL; // OPTION - Hubrahmen oben 303, aus Schaltplan
  Globale_Bausteine.aFaecherwagenstation[303].in_bHubrahmenUnten                                AT %MX1.0    : BOOL; // OPTION - Hubrahmen unten 303, aus Schaltplan
  Globale_Bausteine.aFaecherwagenstation[303].in_bFaecherwagenVorne                             AT %MX1.0    : BOOL; // OPTION - Faecherwagen vorne 303, aus Schaltplan
  Globale_Bausteine.aFaecherwagenstation[303].in_bFaecherwagenHinten                            AT %MX1.0    : BOOL; // OPTION - Faecherwagen hinten 303, aus Schaltplan
  Globale_Bausteine.aFaecherwagenstation[303].in_bZentrierungOffen                              AT %MX1.0    : BOOL; // OPTION - Zentrierung offen 303, aus Schaltplan
  Globale_Bausteine.aFaecherwagenstation[303].in_bZentrierungGeschlossen                        AT %MX1.0    : BOOL; // OPTION - Zentrierung geschlossen 303, aus Schaltplan
  Globale_Bausteine.aFaecherwagenstation[303].in_bAnschlagOben                                  AT %MX1.0    : BOOL; // OPTION - Anschlag oben 303, aus Schaltplan
  Globale_Bausteine.aFaecherwagenstation[303].in_bAnschlagUnten                                 AT %MX1.0    : BOOL; // OPTION - Anschlag unten 303, aus Schaltplan
  Globale_Bausteine.aFaecherwagenstation[303].in_bAnschlagVorne                                 AT %MX1.0    : BOOL; // OPTION - OPTION AGV: Anschlag vorne 303, aus Schaltplan
  Globale_Bausteine.aFaecherwagenstation[303].in_bAnschlagHinten                                AT %MX1.0    : BOOL; // OPTION - OPTION AGV: Anschlag hinten 303, aus Schaltplan
  Globale_Bausteine.aFaecherwagenstation[303].in_bFWInAusrichtPosition                          AT %MX1.0    : BOOL; // OPTION - Faecherwagen in Ausrichtposition 303, aus Schaltplan
  Globale_Bausteine.aFaecherwagenstation[303].in_bMutingSensorLinks                             AT %MX1.0    : BOOL; // OPTION - Muting-Sensor links 303, aus Schaltplan
  Globale_Bausteine.aFaecherwagenstation[303].in_bMutingSensorRechts                            AT %MX1.0    : BOOL; // OPTION - Muting-Sensor rechts 303, aus Schaltplan
  Globale_Bausteine.aFaecherwagenstation[303].in_bStartSchleusen                                AT %MX1.0    : BOOL; // OPTION - Taster Ein-/Ausschleusen 303, aus Schaltplan
  Globale_Bausteine.aFaecherwagenstation[303].in_bSicherheitsrelaisOK                           AT %MX1.1    : BOOL; // OPTION - Sicherheitsrelais in Ordnung 303, aus Schaltplan
  Globale_Bausteine.aFaecherwagenstation[303].in_bAbrollsicherungOK                             AT %MX1.1    : BOOL; // OPTION - Abrollsicherung des Rolltors nicht ausgeloest 303, aus Schaltplan
  Globale_Bausteine.aFaecherwagenstation[303].in_bRFID_DataValid                                AT %MX1.0    : BOOL; // OPTION - RFID Daten gueltig 303, aus Schaltplan
  Globale_Bausteine.aFaecherwagenstation[303].in_bRFID_NR1                                      AT %MX1.0    : BOOL; // OPTION - RFID Bit 1 303, aus Schaltplan
  Globale_Bausteine.aFaecherwagenstation[303].in_bRFID_NR2                                      AT %MX1.0    : BOOL; // OPTION - RFID Bit 2 303, aus Schaltplan
  Globale_Bausteine.aFaecherwagenstation[303].in_bRFID_NR3                                      AT %MX1.0    : BOOL; // OPTION - RFID Bit 3 303, aus Schaltplan
  Globale_Bausteine.aFaecherwagenstation[303].in_bRFID_NR4                                      AT %MX1.0    : BOOL; // OPTION - RFID Bit 4 303, aus Schaltplan
  Globale_Bausteine.aFaecherwagenstation[303].in_bRFID_NR5                                      AT %MX1.0    : BOOL; // OPTION - RFID Bit 5 303, aus Schaltplan
  Globale_Bausteine.aFaecherwagenstation[303].in_bRFID_NR6                                      AT %MX1.0    : BOOL; // OPTION - RFID Bit 6 303, aus Schaltplan
  Globale_Bausteine.aFaecherwagenstation[303].in_bRFID_NR7                                      AT %MX1.0    : BOOL; // OPTION - RFID Bit 7 303, aus Schaltplan
  Globale_Bausteine.aFaecherwagenstation[303].in_bRFID_NR8                                      AT %MX1.0    : BOOL; // OPTION - RFID Bit 8 303, aus Schaltplan
  // AUSGAENGE
  Globale_Bausteine.aFaecherwagenstation[303].out_bHubrahmenHeben                               AT %MX3030.0 : BOOL; // OPTION - Hubrahmen heben 303, aus Schaltplan
  Globale_Bausteine.aFaecherwagenstation[303].out_bHubrahmenSenken                              AT %MX3030.1 : BOOL; // OPTION - Hubrahmen senken 303, aus Schaltplan
  Globale_Bausteine.aFaecherwagenstation[303].out_bFaecherwagenVor                              AT %MX3030.2 : BOOL; // OPTION - Faecherwagen vor 303, aus Schaltplan
  Globale_Bausteine.aFaecherwagenstation[303].out_bFaecherwagenZurueck                          AT %MX3030.3 : BOOL; // OPTION - Faecherwagen zurueck 303, aus Schaltplan
  Globale_Bausteine.aFaecherwagenstation[303].out_bZentrierungOeffnen                           AT %MX3030.4 : BOOL; // OPTION - Zentrierung oeffnen 303, aus Schaltplan
  Globale_Bausteine.aFaecherwagenstation[303].out_bZentrierungSchliessen                        AT %MX3030.5 : BOOL; // OPTION - Zentrierung schliessen 303, aus Schaltplan
  Globale_Bausteine.aFaecherwagenstation[303].out_bAnschlagAuf                                  AT %MX3030.6 : BOOL; // OPTION - Anschlag auf 303, aus Schaltplan
  Globale_Bausteine.aFaecherwagenstation[303].out_bAnschlagAb                                   AT %MX3030.7 : BOOL; // OPTION - Anschlag ab 303, aus Schaltplan
  Globale_Bausteine.aFaecherwagenstation[303].out_bAnschlagVor                                  AT %MX3031.0 : BOOL; // OPTION - OPTION AGV: Anschlag vor 303, aus Schaltplan
  Globale_Bausteine.aFaecherwagenstation[303].out_bAnschlagZurueck                              AT %MX3031.1 : BOOL; // OPTION - OPTION AGV: Anschlag zurueck 303, aus Schaltplan
  Globale_Bausteine.aFaecherwagenstation[303].out_bFreigabeSchleusen                            AT %MX3031.2 : BOOL; // OPTION - Leuchte im Taster Ein-/Ausschleusen 303, aus Schaltplan
  Globale_Bausteine.aFaecherwagenstation[303].out_bMutingSensorReset                            AT %MX3031.3 : BOOL; // OPTION - Reset Muting-Sensoren 303, aus Schaltplan
  Globale_Bausteine.aFaecherwagenstation[303].out_bResetSicherheitsrelais                       AT %MX3031.4 : BOOL; // OPTION - Reset Sicherheitsrelais 303, aus Schaltplan

  // ------------------------------------ STATION 304 ------------------------------------------------
  // EINGAENGE
  Globale_Bausteine.aFaecherwagenstation[304].in_bHubrahmenOben                                 AT %MX1.0    : BOOL; // OPTION - Hubrahmen oben 304, aus Schaltplan
  Globale_Bausteine.aFaecherwagenstation[304].in_bHubrahmenUnten                                AT %MX1.0    : BOOL; // OPTION - Hubrahmen unten 304, aus Schaltplan
  Globale_Bausteine.aFaecherwagenstation[304].in_bFaecherwagenVorne                             AT %MX1.0    : BOOL; // OPTION - Faecherwagen vorne 304, aus Schaltplan
  Globale_Bausteine.aFaecherwagenstation[304].in_bFaecherwagenHinten                            AT %MX1.0    : BOOL; // OPTION - Faecherwagen hinten 304, aus Schaltplan
  Globale_Bausteine.aFaecherwagenstation[304].in_bZentrierungOffen                              AT %MX1.0    : BOOL; // OPTION - Zentrierung offen 304, aus Schaltplan
  Globale_Bausteine.aFaecherwagenstation[304].in_bZentrierungGeschlossen                        AT %MX1.0    : BOOL; // OPTION - Zentrierung geschlossen 304, aus Schaltplan
  Globale_Bausteine.aFaecherwagenstation[304].in_bAnschlagOben                                  AT %MX1.0    : BOOL; // OPTION - Anschlag oben 304, aus Schaltplan
  Globale_Bausteine.aFaecherwagenstation[304].in_bAnschlagUnten                                 AT %MX1.0    : BOOL; // OPTION - Anschlag unten 304, aus Schaltplan
  Globale_Bausteine.aFaecherwagenstation[304].in_bAnschlagVorne                                 AT %MX1.0    : BOOL; // OPTION - OPTION AGV: Anschlag vorne 304, aus Schaltplan
  Globale_Bausteine.aFaecherwagenstation[304].in_bAnschlagHinten                                AT %MX1.0    : BOOL; // OPTION - OPTION AGV: Anschlag hinten 304, aus Schaltplan
  Globale_Bausteine.aFaecherwagenstation[304].in_bFWInAusrichtPosition                          AT %MX1.0    : BOOL; // OPTION - Faecherwagen in Ausrichtposition 304, aus Schaltplan
  Globale_Bausteine.aFaecherwagenstation[304].in_bMutingSensorLinks                             AT %MX1.0    : BOOL; // OPTION - Muting-Sensor links 304, aus Schaltplan
  Globale_Bausteine.aFaecherwagenstation[304].in_bMutingSensorRechts                            AT %MX1.0    : BOOL; // OPTION - Muting-Sensor rechts 304, aus Schaltplan
  Globale_Bausteine.aFaecherwagenstation[304].in_bStartSchleusen                                AT %MX1.0    : BOOL; // OPTION - Taster Ein-/Ausschleusen 304, aus Schaltplan
  Globale_Bausteine.aFaecherwagenstation[304].in_bSicherheitsrelaisOK                           AT %MX1.1    : BOOL; // OPTION - Sicherheitsrelais in Ordnung 304, aus Schaltplan
  Globale_Bausteine.aFaecherwagenstation[304].in_bAbrollsicherungOK                             AT %MX1.1    : BOOL; // OPTION - Abrollsicherung des Rolltors nicht ausgeloest 304, aus Schaltplan
  Globale_Bausteine.aFaecherwagenstation[304].in_bRFID_DataValid                                AT %MX1.0    : BOOL; // OPTION - RFID Daten gueltig 304, aus Schaltplan
  Globale_Bausteine.aFaecherwagenstation[304].in_bRFID_NR1                                      AT %MX1.0    : BOOL; // OPTION - RFID Bit 1 304, aus Schaltplan
  Globale_Bausteine.aFaecherwagenstation[304].in_bRFID_NR2                                      AT %MX1.0    : BOOL; // OPTION - RFID Bit 2 304, aus Schaltplan
  Globale_Bausteine.aFaecherwagenstation[304].in_bRFID_NR3                                      AT %MX1.0    : BOOL; // OPTION - RFID Bit 3 304, aus Schaltplan
  Globale_Bausteine.aFaecherwagenstation[304].in_bRFID_NR4                                      AT %MX1.0    : BOOL; // OPTION - RFID Bit 4 304, aus Schaltplan
  Globale_Bausteine.aFaecherwagenstation[304].in_bRFID_NR5                                      AT %MX1.0    : BOOL; // OPTION - RFID Bit 5 304, aus Schaltplan
  Globale_Bausteine.aFaecherwagenstation[304].in_bRFID_NR6                                      AT %MX1.0    : BOOL; // OPTION - RFID Bit 6 304, aus Schaltplan
  Globale_Bausteine.aFaecherwagenstation[304].in_bRFID_NR7                                      AT %MX1.0    : BOOL; // OPTION - RFID Bit 7 304, aus Schaltplan
  Globale_Bausteine.aFaecherwagenstation[304].in_bRFID_NR8                                      AT %MX1.0    : BOOL; // OPTION - RFID Bit 8 304, aus Schaltplan
  // AUSGAENGE
  Globale_Bausteine.aFaecherwagenstation[304].out_bHubrahmenHeben                               AT %MX3040.0 : BOOL; // OPTION - Hubrahmen heben 304, aus Schaltplan
  Globale_Bausteine.aFaecherwagenstation[304].out_bHubrahmenSenken                              AT %MX3040.1 : BOOL; // OPTION - Hubrahmen senken 304, aus Schaltplan
  Globale_Bausteine.aFaecherwagenstation[304].out_bFaecherwagenVor                              AT %MX3040.2 : BOOL; // OPTION - Faecherwagen vor 304, aus Schaltplan
  Globale_Bausteine.aFaecherwagenstation[304].out_bFaecherwagenZurueck                          AT %MX3040.3 : BOOL; // OPTION - Faecherwagen zurueck 304, aus Schaltplan
  Globale_Bausteine.aFaecherwagenstation[304].out_bZentrierungOeffnen                           AT %MX3040.4 : BOOL; // OPTION - Zentrierung oeffnen 304, aus Schaltplan
  Globale_Bausteine.aFaecherwagenstation[304].out_bZentrierungSchliessen                        AT %MX3040.5 : BOOL; // OPTION - Zentrierung schliessen 304, aus Schaltplan
  Globale_Bausteine.aFaecherwagenstation[304].out_bAnschlagAuf                                  AT %MX3040.6 : BOOL; // OPTION - Anschlag auf 304, aus Schaltplan
  Globale_Bausteine.aFaecherwagenstation[304].out_bAnschlagAb                                   AT %MX3040.7 : BOOL; // OPTION - Anschlag ab 304, aus Schaltplan
  Globale_Bausteine.aFaecherwagenstation[304].out_bAnschlagVor                                  AT %MX3041.0 : BOOL; // OPTION - OPTION AGV: Anschlag vor 304, aus Schaltplan
  Globale_Bausteine.aFaecherwagenstation[304].out_bAnschlagZurueck                              AT %MX3041.1 : BOOL; // OPTION - OPTION AGV: Anschlag zurueck 304, aus Schaltplan
  Globale_Bausteine.aFaecherwagenstation[304].out_bFreigabeSchleusen                            AT %MX3041.2 : BOOL; // OPTION - Leuchte im Taster Ein-/Ausschleusen 304, aus Schaltplan
  Globale_Bausteine.aFaecherwagenstation[304].out_bMutingSensorReset                            AT %MX3041.3 : BOOL; // OPTION - Reset Muting-Sensoren 304, aus Schaltplan
  Globale_Bausteine.aFaecherwagenstation[304].out_bResetSicherheitsrelais                       AT %MX3041.4 : BOOL; // OPTION - Reset Sicherheitsrelais 304, aus Schaltplan

  // ------------------------------------ STATION 305 ------------------------------------------------
  // EINGAENGE
  Globale_Bausteine.aFaecherwagenstation[305].in_bHubrahmenOben                                 AT %MX1.0    : BOOL; // OPTION - Hubrahmen oben 305, aus Schaltplan
  Globale_Bausteine.aFaecherwagenstation[305].in_bHubrahmenUnten                                AT %MX1.0    : BOOL; // OPTION - Hubrahmen unten 305, aus Schaltplan
  Globale_Bausteine.aFaecherwagenstation[305].in_bFaecherwagenVorne                             AT %MX1.0    : BOOL; // OPTION - Faecherwagen vorne 305, aus Schaltplan
  Globale_Bausteine.aFaecherwagenstation[305].in_bFaecherwagenHinten                            AT %MX1.0    : BOOL; // OPTION - Faecherwagen hinten 305, aus Schaltplan
  Globale_Bausteine.aFaecherwagenstation[305].in_bZentrierungOffen                              AT %MX1.0    : BOOL; // OPTION - Zentrierung offen 305, aus Schaltplan
  Globale_Bausteine.aFaecherwagenstation[305].in_bZentrierungGeschlossen                        AT %MX1.0    : BOOL; // OPTION - Zentrierung geschlossen 305, aus Schaltplan
  Globale_Bausteine.aFaecherwagenstation[305].in_bAnschlagOben                                  AT %MX1.0    : BOOL; // OPTION - Anschlag oben 305, aus Schaltplan
  Globale_Bausteine.aFaecherwagenstation[305].in_bAnschlagUnten                                 AT %MX1.0    : BOOL; // OPTION - Anschlag unten 305, aus Schaltplan
  Globale_Bausteine.aFaecherwagenstation[305].in_bAnschlagVorne                                 AT %MX1.0    : BOOL; // OPTION - OPTION AGV: Anschlag vorne 305, aus Schaltplan
  Globale_Bausteine.aFaecherwagenstation[305].in_bAnschlagHinten                                AT %MX1.0    : BOOL; // OPTION - OPTION AGV: Anschlag hinten 305, aus Schaltplan
  Globale_Bausteine.aFaecherwagenstation[305].in_bFWInAusrichtPosition                          AT %MX1.0    : BOOL; // OPTION - Faecherwagen in Ausrichtposition 305, aus Schaltplan
  Globale_Bausteine.aFaecherwagenstation[305].in_bMutingSensorLinks                             AT %MX1.0    : BOOL; // OPTION - Muting-Sensor links 305, aus Schaltplan
  Globale_Bausteine.aFaecherwagenstation[305].in_bMutingSensorRechts                            AT %MX1.0    : BOOL; // OPTION - Muting-Sensor rechts 305, aus Schaltplan
  Globale_Bausteine.aFaecherwagenstation[305].in_bStartSchleusen                                AT %MX1.0    : BOOL; // OPTION - Taster Ein-/Ausschleusen 305, aus Schaltplan
  Globale_Bausteine.aFaecherwagenstation[305].in_bSicherheitsrelaisOK                           AT %MX1.1    : BOOL; // OPTION - Sicherheitsrelais in Ordnung 305, aus Schaltplan
  Globale_Bausteine.aFaecherwagenstation[305].in_bAbrollsicherungOK                             AT %MX1.1    : BOOL; // OPTION - Abrollsicherung des Rolltors nicht ausgeloest 305, aus Schaltplan
  Globale_Bausteine.aFaecherwagenstation[305].in_bRFID_DataValid                                AT %MX1.0    : BOOL; // OPTION - RFID Daten gueltig 305, aus Schaltplan
  Globale_Bausteine.aFaecherwagenstation[305].in_bRFID_NR1                                      AT %MX1.0    : BOOL; // OPTION - RFID Bit 1 305, aus Schaltplan
  Globale_Bausteine.aFaecherwagenstation[305].in_bRFID_NR2                                      AT %MX1.0    : BOOL; // OPTION - RFID Bit 2 305, aus Schaltplan
  Globale_Bausteine.aFaecherwagenstation[305].in_bRFID_NR3                                      AT %MX1.0    : BOOL; // OPTION - RFID Bit 3 305, aus Schaltplan
  Globale_Bausteine.aFaecherwagenstation[305].in_bRFID_NR4                                      AT %MX1.0    : BOOL; // OPTION - RFID Bit 4 305, aus Schaltplan
  Globale_Bausteine.aFaecherwagenstation[305].in_bRFID_NR5                                      AT %MX1.0    : BOOL; // OPTION - RFID Bit 5 305, aus Schaltplan
  Globale_Bausteine.aFaecherwagenstation[305].in_bRFID_NR6                                      AT %MX1.0    : BOOL; // OPTION - RFID Bit 6 305, aus Schaltplan
  Globale_Bausteine.aFaecherwagenstation[305].in_bRFID_NR7                                      AT %MX1.0    : BOOL; // OPTION - RFID Bit 7 305, aus Schaltplan
  Globale_Bausteine.aFaecherwagenstation[305].in_bRFID_NR8                                      AT %MX1.0    : BOOL; // OPTION - RFID Bit 8 305, aus Schaltplan
  // AUSGAENGE
  Globale_Bausteine.aFaecherwagenstation[305].out_bHubrahmenHeben                               AT %MX3050.0 : BOOL; // OPTION - Hubrahmen heben 305, aus Schaltplan
  Globale_Bausteine.aFaecherwagenstation[305].out_bHubrahmenSenken                              AT %MX3050.1 : BOOL; // OPTION - Hubrahmen senken 305, aus Schaltplan
  Globale_Bausteine.aFaecherwagenstation[305].out_bFaecherwagenVor                              AT %MX3050.2 : BOOL; // OPTION - Faecherwagen vor 305, aus Schaltplan
  Globale_Bausteine.aFaecherwagenstation[305].out_bFaecherwagenZurueck                          AT %MX3050.3 : BOOL; // OPTION - Faecherwagen zurueck 305, aus Schaltplan
  Globale_Bausteine.aFaecherwagenstation[305].out_bZentrierungOeffnen                           AT %MX3050.4 : BOOL; // OPTION - Zentrierung oeffnen 305, aus Schaltplan
  Globale_Bausteine.aFaecherwagenstation[305].out_bZentrierungSchliessen                        AT %MX3050.5 : BOOL; // OPTION - Zentrierung schliessen 305, aus Schaltplan
  Globale_Bausteine.aFaecherwagenstation[305].out_bAnschlagAuf                                  AT %MX3050.6 : BOOL; // OPTION - Anschlag auf 305, aus Schaltplan
  Globale_Bausteine.aFaecherwagenstation[305].out_bAnschlagAb                                   AT %MX3050.7 : BOOL; // OPTION - Anschlag ab 305, aus Schaltplan
  Globale_Bausteine.aFaecherwagenstation[305].out_bAnschlagVor                                  AT %MX3051.0 : BOOL; // OPTION - OPTION AGV: Anschlag vor 305, aus Schaltplan
  Globale_Bausteine.aFaecherwagenstation[305].out_bAnschlagZurueck                              AT %MX3051.1 : BOOL; // OPTION - OPTION AGV: Anschlag zurueck 305, aus Schaltplan
  Globale_Bausteine.aFaecherwagenstation[305].out_bFreigabeSchleusen                            AT %MX3051.2 : BOOL; // OPTION - Leuchte im Taster Ein-/Ausschleusen 305, aus Schaltplan
  Globale_Bausteine.aFaecherwagenstation[305].out_bMutingSensorReset                            AT %MX3051.3 : BOOL; // OPTION - Reset Muting-Sensoren 305, aus Schaltplan
  Globale_Bausteine.aFaecherwagenstation[305].out_bResetSicherheitsrelais                       AT %MX3051.4 : BOOL; // OPTION - Reset Sicherheitsrelais 305, aus Schaltplan

END_VAR

END_NAMESPACE
